Fanuc KAREL source: kb00041.KL

-- PROVISIONAL review KL for V940-1; original PC SHA256 676e73277c41af3ba342b3d420ffcc326a144e4dba9b6f4fdb24b5d17a5429f5
-- Incomplete behavior may be omitted. Consult companion uncertainty JSON. Do not deploy.
PROGRAM KB00041
%NOLOCKGROUP
BEGIN
  -- V9_ZERO_TABLE_METADATA_HINT layout=0002_ascii; no indexed target words; source/name/runtime held
  -- UNRESOLVED_PC offsets 5-14; opcodes 3F,75
  -- UNRESOLVED_PC offsets 19-30; opcodes 2E,23
  -- UNRESOLVED_PC offsets 35-53; opcodes 27,22,2A,22,31
  -- UNRESOLVED_PC offsets 58-62; opcodes 7F
END KB00041
